// TIA Portal V21 export
// export: Created 2026-11-22T00:27:33.9071901Z, ExportSetting WithDefaults, DisplayName Totally Integrated Automation Portal, DisplayVersion V21 Update 3, DisplayName STEP 7 Professional, DisplayVersion V21 Update 3, DisplayName STEP 7 Safety, DisplayVersion V21, DisplayName Tech WebApplication, DisplayVersion V21, DisplayName WinCC Basic/Comfort/Advanced, DisplayVersion V21 Update 3, DisplayName WinCC Unified, DisplayVersion V21 Update 3
Screen "P_Bar_2"  800x480, Number=114
  ScreenLayer "Layer_0"
    Bar "ShowTickLabels" at 10,10 size 40x120  CountSubDivisions=5, IntegerDigits=3, LargeTickLabelingStep=1, MaximumValue=5, MinimumValue=-5, Precision=2, StyleItem=Bar
    TextField "Label_ShowTickLabels" at 10,132 size 48x16  StyleItem=Text field, Text="ShowTickLabels"
    Bar "Unit" at 60,10 size 40x120  CountSubDivisions=5, IntegerDigits=3, LargeTickLabelingStep=1, MaximumValue=5, MinimumValue=-5, Precision=2, Unit=mm, StyleItem=Bar
    TextField "Label_Unit" at 60,132 size 48x16  StyleItem=Text field, Text="Unit"
    Bar "UseAutoScaling" at 110,10 size 40x120  CountSubDivisions=5, IntegerDigits=3, LargeTickLabelingStep=1, MaximumValue=5, MinimumValue=-5, Precision=2, StyleItem=Bar
    TextField "Label_UseAutoScaling" at 110,132 size 48x16  StyleItem=Text field, Text="UseAutoScaling"
    Bar "UseDesignColorSchema" at 160,10 size 40x120  CountSubDivisions=5, IntegerDigits=3, LargeTickLabelingStep=1, MaximumValue=5, MinimumValue=-5, Precision=2
    TextField "Label_UseDesignColorSchema" at 160,132 size 48x16  StyleItem=Text field, Text="UseDesignColorSchema"
    Bar "UseExponentialFormat" at 210,10 size 40x120  CountSubDivisions=5, IntegerDigits=3, LargeTickLabelingStep=1, MaximumValue=5, MinimumValue=-5, Precision=2, StyleItem=Bar
    TextField "Label_UseExponentialFormat" at 210,132 size 48x16  StyleItem=Text field, Text="UseExponentialFormat"
    Button "Next" at 758,456 size 40x22  Mode=Text, StyleItem=Button, TextOff="Text", TextOn="Text"
      on Click: ActivateScreen(Screen name := P_Switch_1, Object number := 0)
